// TIA Portal V21 export
// export: Created 2026-08-21T20:18:56.912201Z, ExportSetting None, DisplayName Totally Integrated Automation Portal, DisplayVersion V21, DisplayName STEP 7 Professional, DisplayVersion V21, DisplayName STEP 7 Safety, DisplayVersion V21, DisplayName Tech WebApplication, DisplayVersion V21, DisplayName WinCC Basic/Comfort/Advanced, DisplayVersion V21, DisplayName WinCC Professional, DisplayVersion V21, DisplayName WinCC Unified, DisplayVersion V21
TYPE "UDT_Service_ParameterDataMedium"
   STRUCT
      used : Array[0..0] of DWord;   // Used configuration parameters of service
      definition : Array[0..31] of "UDT_Service_ParameterDefinition";
   END_STRUCT;
END_TYPE
